(* IEC 61131-3 sources: Elmo_Master/Lasal_PRG/MotionTCPDemo/Class/_SigTCPDataManager, 1 file *)

(* ---- _SigTCPDataManager.st ---- *)
(*!
<Class
	Name               = "_SigTCPDataManager"
	Revision           = "1.1"
	RealtimeTask       = "false"
	CyclicTask         = "true"
	DefCyclictime      = "100 ms"
	BackgroundTask     = "false"
	Sigmatek           = "true"
	OSInterface        = "false"
	HighPriority       = "false"
	Automatic          = "false"
	UpdateMode         = "Prescan"
	SharedCommandTable = "true"
	Objectsize         = "(678,120)"
	Comment            = "This class is designed to simplify the implementation of TCP communication.&#13;&#10;It already contains the TCPCommunication and DataManager classes.&#13;&#10;&#13;&#10;The _SigTCPComSend and _SigTCPComReceive classes can be directly connected and operated with this class.">
	<Channels>
		<Server Name="ComPort" Visualized="true" Initialize="true" WriteProtected="false" Retentive="false" Comment="The TCP Port which is used for communication has to be configured here. &#13;&#10;Sender and Receiver have to use the same port.&#13;&#10;&#13;&#10;If there are multiple senders or receivers in the same project, different ports must be used.&#13;&#10;&#13;&#10;e.g.: Sender1 - Receiver1 -&gt; 500&#13;&#10;       Sender2 - Receiver2 -&gt; 600"/>
		<Server Name="DeactivateCom" Visualized="false" Initialize="true" WriteProtected="false" Retentive="false" Comment="Set to 1 to deactivate communication.&#13;&#10;Set to 0 to reactivate communication."/>
		<Server Name="LogEnable" Visualized="true" Initialize="true" WriteProtected="false" Retentive="false" Comment="0 = Logging is deactivated&#13;&#10;1 = Logging is active"/>
		<Server Name="Online" Visualized="true" Initialize="false" WriteProtected="true" Retentive="false" Comment="State of the connection &#13;&#10;0 = Offline&#13;&#10;1 = Online"/>
		<Server Name="ResetLogBuffer" Visualized="true" Initialize="false" WriteProtected="false" Retentive="false" Comment="Write() on this Server deletes the internal log buffer. &#13;&#10;Can only be executed if the server LogEnable is set to 0."/>
		<Server Name="TCPComm" Class="TCPCommunication" Visualized="true" Initialize="false" WriteProtected="false" Retentive="false" Comment="Object server of the class TCPCommunication. &#13;&#10;Can be used to call the global methods of the TCPCommunication class.&#13;&#10;The class TCPCommunicationLogViewer can be connected to this server in order to read and export the log entries."/>
		<Client Name="ErrRuntime" Required="false" Internal="false" Comment="If the parallel communication task was not called for longer than TCPCom_Runtime (tcpcommunication.h), this Client will turn to 1 and if a Server is connected, it&apos;s write-Method will be called with input:=1.&#13;&#10;If it is called again after that, the Client will turn to 0 again and the write method will be called again with input:=0.&#13;&#10;Also, a TRACE-Error will be caused when the error is detected, and a TRACE-Warning will be caused as soon as the parallel task is running again."/>
		<Client Name="InternConnection" Required="false" Internal="false" Comment="If an external connection (via TCPIP) shall be established, this client may not be connected!&#13;&#10;&#13;&#10;If the connection is internal (sender and receiver are on the same cpu), this client has to be connected to the ClassSvr of the corresponding TCPCommunication class.&#13;&#10;"/>
		<Client Name="IPtoConnect" Required="false" Internal="false" Comment="Required if the class should work as a TCPIP client. &#13;&#10;Connection to an object of the String or StringRAM class &#13;&#10;(IP address of the desired TCPIP server to connect)."/>
		<Client Name="LogFilter" Required="false" Internal="false" Comment="If the TCPCommunicationLogFilter is used, it has to be connected here."/>
		<Client Name="SizeOfComBufferRecv" Required="false" Internal="false" Comment="Size of the receive buffer. Has to be set as Init-Value!&#13;&#10;If the allocated memory is too small for the received buffer the variable dRecvErrorBuffersize shows the needed size."/>
		<Client Name="SizeOfComBuffers" Required="false" Internal="false" Comment="Size of the send buffer. Has to be set as Init-Value!"/>
		<Client Name="StationToConnect" Required="false" Internal="false" Comment="Connect it to class &quot;GetIPOverStation&quot; server &quot;ClassSvr&quot; to get the ip address over set station number."/>
		<Client Name="TCPCommunication" Required="true" Internal="true"/>
	</Channels>
	<Separators>
		<Servers>
			<SepChn Position="0"/>
		</Servers>
	</Separators>
	<RevDoku>
		<Owner Company="Sigmatek"/>
		<Dokumentation Revision="1.1" Date="2025-09-30" Author="KaiAnd" Company="Sigmatek" Description="Optimized comments and style"/>
		<Dokumentation Revision="1.0" Date="2025-04-24" Author="SchMar2" Company="Sigmatek" Description="Initial version"/>
	</RevDoku>
	<Network Name="_SigTCPDataManager">
		<!-- List of Components in this network -->
		<Components>
			<Object
				Name       = "_base"
				Class      = "DataManager"
				Position   = "(1134,150)"
				Visualized = "false">
				<Channels>
					<Server Name="AcceptOfflineJobs" Value="1"/>
					<Server Name="ClassSvr"/>
					<Server Name="DeleteJobs"/>
					<Server Name="NoEntries"/>
					<Client Name="coTCPCommunication"/>
				</Channels>
			</Object>
			<Object
				Name       = "TCPCommunication"
				Class      = "TCPCommunication"
				Position   = "(360,150)"
				Visualized = "false">
				<Channels>
					<Server Name="ClassSvr"/>
					<Server Name="ComPort" Value="500"/>
					<Server Name="ConnectionType"/>
					<Server Name="DeactivateCom" Value="0"/>
					<Server Name="ErrorRecive"/>
					<Server Name="ErrorSend"/>
					<Server Name="InitError"/>
					<Server Name="LogEnable" Value="0"/>
					<Server Name="Online"/>
					<Server Name="ResetLogBuffer"/>
					<Server Name="TaskName"/>
					<Server Name="TimeLastReceive"/>
					<Server Name="TimeLastSend"/>
					<Server Name="TransferRateReceive"/>
					<Server Name="TransferRateSend"/>
					<Client Name="coDataMng"/>
					<Client Name="coIntern"/>
					<Client Name="coIpToConnect"/>
					<Client Name="coLogFilter" Value="0"/>
					<Client Name="coMultiTask"/>
					<Client Name="coSigCLib"/>
					<Client Name="coStationToConnect"/>
					<Client Name="coStdLib"/>
					<Client Name="ErrRuntime"/>
					<Client Name="SizeOfComBufferRecv" Value="100 kB"/>
					<Client Name="SizeOfComBuffers" Value="100 kB"/>
				</Channels>
			</Object>
		</Components>
		<Comments>
		</Comments>
		<!-- List of Connections in this network -->
		<Connections>
			<Connection Source="this.TCPCommunication" Destination="TCPCommunication.ClassSvr"/>
			<Connection Source="_base.coTCPCommunication" Destination="TCPCommunication.ClassSvr" Vertices="(1134,240),(1008,240),"/>
			<Connection Source="TCPCommunication.coDataMng" Destination="_base.ClassSvr" Vertices="(360,240),(330,240),(330,120),(1860,120),(1860,240),(1810,240),"/>
			<Connection Source="this.LogEnable" Destination="TCPCommunication.LogEnable" Vertices="(1982,630),(1008,900),"/>
			<Connection Source="TCPCommunication.coIntern" Destination="this.InternConnection" Vertices="(360,300),(38,450),"/>
			<Connection Source="this.ClassSvr" Destination="_base.ClassSvr" Vertices="(1982,210),(1810,240),"/>
			<Connection Source="this.NoEntries" Destination="_base.NoEntries" Vertices="(1982,270),(1810,300),"/>
			<Connection Source="this.DeleteJobs" Destination="_base.DeleteJobs" Vertices="(1982,330),(1810,360),"/>
			<Connection Source="TCPCommunication.coIpToConnect" Destination="this.IPtoConnect" Vertices="(360,360),(38,510),"/>
			<Connection Source="TCPCommunication.coStationToConnect" Destination="this.StationToConnect" Vertices="(360,420),(38,570),"/>
			<Connection Source="TCPCommunication.coLogFilter" Destination="this.LogFilter" Vertices="(360,480),(38,630),"/>
			<Connection Source="TCPCommunication.ErrRuntime" Destination="this.ErrRuntime" Vertices="(360,720),(38,690),"/>
			<Connection Source="TCPCommunication.SizeOfComBuffers" Destination="this.SizeOfComBuffers" Vertices="(360,780),(38,750),"/>
			<Connection Source="TCPCommunication.SizeOfComBufferRecv" Destination="this.SizeOfComBufferRecv" Vertices="(360,840),(38,810),"/>
			<Connection Source="this.AcceptOfflineJobs" Destination="_base.AcceptOfflineJobs" Vertices="(1982,390),(1810,420),"/>
			<Connection Source="this.ResetLogBuffer" Destination="TCPCommunication.ResetLogBuffer" Vertices="(1982,690),(1008,960),"/>
			<Connection Source="this.ComPort" Destination="TCPCommunication.ComPort" Vertices="(1982,510),(1008,420),"/>
			<Connection Source="this.Online" Destination="TCPCommunication.Online" Vertices="(1982,570),(1290,510),(1008,480),"/>
			<Connection Source="this.DeactivateCom" Destination="TCPCommunication.DeactivateCom" Vertices="(1982,750),(1008,1080),"/>
			<Connection Source="this.TCPComm" Destination="TCPCommunication.ClassSvr" Vertices="(1982,450),(1008,240),"/>
		</Connections>
		<!-- Headerfiles -->
		<Options>
		</Options>
	</Network>
</Class>
*)
#pragma using DataManager

_SigTCPDataManager : CLASS
: DataManager
  //Servers:
	TCPComm 	: SvrChCmd_DINT;
	ComPort 	: SvrCh_UDINT;
	Online 	: SvrCh_DINT;
	LogEnable 	: SvrCh_DINT;
	ResetLogBuffer 	: SvrCh_DINT;
	DeactivateCom 	: SvrCh_DINT;
  //Clients:
	TCPCommunication 	: CltChCmd_TCPCommunication;
	InternConnection 	: CltChCmd_TCPCommunication;
	IPtoConnect 	: CltChCmd_StringInternal;
	StationToConnect 	: CltChCmd_DINT;
	LogFilter 	: CltChCmd_TCPCommunicationLogFilter;
	ErrRuntime 	: CltCh_DINT;
	SizeOfComBuffers 	: CltCh_UDINT;
	SizeOfComBufferRecv 	: CltCh_UDINT;
  //Variables:
  //Functions:
				//! <Function Comment="Cyclic Work" Name="CyWork"/>
	FUNCTION VIRTUAL GLOBAL CyWork
		VAR_INPUT
			EAX 	: UDINT;
		END_VAR
		VAR_OUTPUT
			state (EAX) 	: UDINT;
		END_VAR;

	FUNCTION VIRTUAL GLOBAL TCPComm::Read
		VAR_OUTPUT
			output (EAX) 	: DINT;
		END_VAR;

	FUNCTION VIRTUAL GLOBAL TCPComm::Write
		VAR_INPUT
			input (EAX) 	: DINT;
		END_VAR
		VAR_OUTPUT
			result (EAX) 	: DINT;
		END_VAR;

	FUNCTION VIRTUAL GLOBAL ComPort::Read
		VAR_OUTPUT
			output (EAX) 	: UDINT;
		END_VAR;

	FUNCTION VIRTUAL GLOBAL ComPort::Write
		VAR_INPUT
			input (EAX) 	: UDINT;
		END_VAR
		VAR_OUTPUT
			result (EAX) 	: UDINT;
		END_VAR;

	FUNCTION VIRTUAL GLOBAL Online::Read
		VAR_OUTPUT
			output (EAX) 	: DINT;
		END_VAR;

	FUNCTION VIRTUAL GLOBAL LogEnable::Read
		VAR_OUTPUT
			output (EAX) 	: DINT;
		END_VAR;

	FUNCTION VIRTUAL GLOBAL LogEnable::Write
		VAR_INPUT
			input (EAX) 	: DINT;
		END_VAR
		VAR_OUTPUT
			result (EAX) 	: DINT;
		END_VAR;

	FUNCTION VIRTUAL GLOBAL ResetLogBuffer::Read
		VAR_OUTPUT
			output (EAX) 	: DINT;
		END_VAR;

	FUNCTION VIRTUAL GLOBAL ResetLogBuffer::Write
		VAR_INPUT
			input (EAX) 	: DINT;
		END_VAR
		VAR_OUTPUT
			result (EAX) 	: DINT;
		END_VAR;

	FUNCTION VIRTUAL GLOBAL DeactivateCom::Read
		VAR_OUTPUT
			output (EAX) 	: DINT;
		END_VAR;

	FUNCTION VIRTUAL GLOBAL DeactivateCom::Write
		VAR_INPUT
			input (EAX) 	: DINT;
		END_VAR
		VAR_OUTPUT
			result (EAX) 	: DINT;
		END_VAR;
  //Tables:
	FUNCTION @STD
		VAR_OUTPUT
			ret_code	: CONFSTATES;
		END_VAR;
	FUNCTION GLOBAL TAB @CT_;
END_CLASS;

#pragma using TCPCommunication
#pragma usingLtd StringInternal
#pragma usingLtd TCPCommunicationLogFilter

FUNCTION VIRTUAL GLOBAL _SigTCPDataManager::CyWork
	VAR_INPUT
		EAX 	: UDINT;
	END_VAR
	VAR_OUTPUT
		state (EAX) 	: UDINT;
	END_VAR

  // call cywork of tcp communication so no task settings need to be done in complex network
  TCPCommunication.CyWork(EAX);

	state := READY;

END_FUNCTION

FUNCTION VIRTUAL GLOBAL _SigTCPDataManager::TCPComm::Read
	VAR_OUTPUT
		output (EAX) 	: DINT;
	END_VAR

	TCPComm := TCPCommunication.ClassSvr.Read();
	output := TCPComm;

END_FUNCTION

FUNCTION VIRTUAL GLOBAL _SigTCPDataManager::TCPComm::Write
	VAR_INPUT
		input (EAX) 	: DINT;
	END_VAR
	VAR_OUTPUT
		result (EAX) 	: DINT;
	END_VAR

	TCPComm := input;
	result := (TCPCommunication.ClassSvr.Write(TCPComm))$DINT;

END_FUNCTION

FUNCTION VIRTUAL GLOBAL _SigTCPDataManager::ComPort::Read
	VAR_OUTPUT
		output (EAX) 	: UDINT;
	END_VAR

	ComPort := TCPCommunication.ComPort.Read();
	output := ComPort;

END_FUNCTION

FUNCTION VIRTUAL GLOBAL _SigTCPDataManager::ComPort::Write
	VAR_INPUT
		input (EAX) 	: UDINT;
	END_VAR
	VAR_OUTPUT
		result (EAX) 	: UDINT;
	END_VAR

	ComPort := input;
	result := (TCPCommunication.ComPort.Write(ComPort))$UDINT;

END_FUNCTION

FUNCTION VIRTUAL GLOBAL _SigTCPDataManager::Online::Read
	VAR_OUTPUT
		output (EAX) 	: DINT;
	END_VAR

	Online := TCPCommunication.Online.Read();
	output := Online;

END_FUNCTION

FUNCTION VIRTUAL GLOBAL _SigTCPDataManager::LogEnable::Read
	VAR_OUTPUT
		output (EAX) 	: DINT;
	END_VAR

	LogEnable := TCPCommunication.LogEnable.Read();
	output := LogEnable;

END_FUNCTION

FUNCTION VIRTUAL GLOBAL _SigTCPDataManager::LogEnable::Write
	VAR_INPUT
		input (EAX) 	: DINT;
	END_VAR
	VAR_OUTPUT
		result (EAX) 	: DINT;
	END_VAR

	LogEnable := input;
	result := (TCPCommunication.LogEnable.Write(LogEnable))$DINT;

END_FUNCTION

FUNCTION VIRTUAL GLOBAL _SigTCPDataManager::ResetLogBuffer::Read
	VAR_OUTPUT
		output (EAX) 	: DINT;
	END_VAR

	ResetLogBuffer := TCPCommunication.ResetLogBuffer.Read();
	output := ResetLogBuffer;

END_FUNCTION

FUNCTION VIRTUAL GLOBAL _SigTCPDataManager::ResetLogBuffer::Write
	VAR_INPUT
		input (EAX) 	: DINT;
	END_VAR
	VAR_OUTPUT
		result (EAX) 	: DINT;
	END_VAR

	ResetLogBuffer := input;
	result := (TCPCommunication.ResetLogBuffer.Write(ResetLogBuffer))$DINT;

END_FUNCTION

FUNCTION VIRTUAL GLOBAL _SigTCPDataManager::DeactivateCom::Read
	VAR_OUTPUT
		output (EAX) 	: DINT;
	END_VAR

	DeactivateCom := TCPCommunication.DeactivateCom.Read();
	output := DeactivateCom;

END_FUNCTION

FUNCTION VIRTUAL GLOBAL _SigTCPDataManager::DeactivateCom::Write
	VAR_INPUT
		input (EAX) 	: DINT;
	END_VAR
	VAR_OUTPUT
		result (EAX) 	: DINT;
	END_VAR

	DeactivateCom := input;
	result := (TCPCommunication.DeactivateCom.Write(DeactivateCom))$DINT;

END_FUNCTION
